PROGRAM MAIN
VAR
	fb : FB_MainControlCell; 
	fb1 : FB_StationBase;
END_VAR

END_PROGRAM

(* stored: Version 1.1.0.1, ProductVersion 3.1.4024.12
   POU MAIN: Id {d1cc440d-f64c-4812-8b56-54077dbf711b}, SpecialFunc None *)
